// TIA Portal V20 export
VAR_GLOBAL   // PLC tag table "laser_out_macsa"
   "-XT500_output_mode" AT %QD295 : DWord;   // Pole - výber pole podle čísla max 255
   "-XT500_output_byte_1" AT %QB295 : Byte;
   "-XT500_output_byte_2" AT %QB296 : Byte;
   "-XT500_output_byte_3" AT %QB297 : Byte;
   "-XT500_output_byte_4" AT %QB298 : Byte;
   "-XT500_output_copies" AT %QD299 : DWord;
   "-XT500_output_byte_5" AT %QB299 : Byte;   // zapisovaná data
   "-XT500_output_byte_6" AT %QB300 : Byte;   // zapisovaná data
   "-XT500_output_byte_7" AT %QB301 : Byte;   // zapisovaná data
   "-XT500_output_byte_8" AT %QB302 : Byte;   // zapisovaná data
   "-XT500_output_byte_9" AT %QB303 : Byte;   // zapisovaná data
   "-XT500_output_batch" AT %QD303 : DWord;
   "-XT500_output_byte_10" AT %QB304 : Byte;   // zapisovaná data
   "-XT500_output_byte_11" AT %QB305 : Byte;   // zapisovaná data
   "-XT500_output_byte_12" AT %QB306 : Byte;   // zapisovaná data
   "-XT500_output_filename_1" AT %QB307 : Byte;   // zápid textu v asci pro volbu programu + další data
   "-XT500_output_filename_2" AT %QB308 : Byte;   // zápid textu v asci pro volbu programu + další data
   "-XT500_output_filename_3" AT %QB309 : Byte;   // zápid textu v asci pro volbu programu + další data
   "-XT500_output_filename_4" AT %QB310 : Byte;   // zápid textu v asci pro volbu programu + další data
   "-XT500_output_filename_5" AT %QB311 : Byte;   // zápid textu v asci pro volbu programu + další data
   "-XT500_output_filename_6" AT %QB312 : Byte;   // zápid textu v asci pro volbu programu + další data
   "-XT500_output_filename_7" AT %QB313 : Byte;   // zápid textu v asci pro volbu programu + další data
   "-XT500_output_filename_8" AT %QB314 : Byte;   // zápid textu v asci pro volbu programu + další data
   "-XT500_output_filename_9" AT %QB315 : Byte;   // zápid textu v asci pro volbu programu + další data
   "-XT500_output_filename_10" AT %QB316 : Byte;   // zápid textu v asci pro volbu programu + další data
   "-XT500_output_filename_11" AT %QB317 : Byte;   // zápid textu v asci pro volbu programu + další data
   "-XT500_output_filename_12" AT %QB318 : Byte;   // zápid textu v asci pro volbu programu + další data
   "-XT500_output_filename_13" AT %QB319 : Byte;   // zápid textu v asci pro volbu programu + další data
   "-XT500_output_filename_14" AT %QB320 : Byte;   // zápid textu v asci pro volbu programu + další data
   "-XT500_output_filename_15" AT %QB321 : Byte;   // zápid textu v asci pro volbu programu + další data
   "-XT500_output_filename_16" AT %QB322 : Byte;   // zápid textu v asci pro volbu programu + další data
   "-XT500_output_filename_17" AT %QB323 : Byte;   // zápid textu v asci pro volbu programu + další data
   "-XT500_command_number" AT %QB293 : Byte;   // výběr daného komandu v podobě čísla podle návodu zadavano v decu pozor na převod mezi word a int ----------- 6 zapis dat 16 vypal 1 otevření zprávy
   "-XT500_command_triger" AT %QB294 : Byte;   // 1= proveď příkaz
   "-XT500_output_filename_18" AT %QB324 : Byte;   // zápid textu v asci pro volbu programu + další data
   "-XT500_output_filename_19" AT %QB325 : Byte;   // zápid textu v asci pro volbu programu + další data
   "-XT500_output_filename_20" AT %QB326 : Byte;   // zápid textu v asci pro volbu programu + další data
   "-XT500_output_filename_21" AT %QB327 : Byte;   // zápid textu v asci pro volbu programu + další data
   "-XT500_output_filename_22" AT %QB328 : Byte;   // zápid textu v asci pro volbu programu + další data
   "-XT500_output_filename_23" AT %QB329 : Byte;   // zápid textu v asci pro volbu programu + další data
   "-XT500_output_filename_24" AT %QB330 : Byte;   // zápid textu v asci pro volbu programu + další data
   "-XT500_output_filename_25" AT %QB331 : Byte;   // zápid textu v asci pro volbu programu + další data
   "-XT500_output_filename_26" AT %QB332 : Byte;   // zápid textu v asci pro volbu programu + další data
   "-XT500_output_filename_27" AT %QB333 : Byte;   // zápid textu v asci pro volbu programu + další data
   "-XT500_output_filename_28" AT %QB334 : Byte;   // zápid textu v asci pro volbu programu + další data
   "-XT500_output_filename_29" AT %QB335 : Byte;   // zápid textu v asci pro volbu programu + další data
   "-XT500_output_filename_30" AT %QB336 : Byte;   // zápid textu v asci pro volbu programu + další data
   "-XT500_output_filename_31" AT %QB337 : Byte;   // zápid textu v asci pro volbu programu + další data
   "-XT500_output_filename_32" AT %QB338 : Byte;   // zápid textu v asci pro volbu programu + další data
   "-XT500_output_filename_33" AT %QB339 : Byte;   // zápid textu v asci pro volbu programu + další data
   "-XT500_output_filename_34" AT %QB340 : Byte;   // zápid textu v asci pro volbu programu + další data
   "-XT500_output_filename_35" AT %QB341 : Byte;   // zápid textu v asci pro volbu programu + další data
   "-XT500_output_filename_36" AT %QB342 : Byte;   // zápid textu v asci pro volbu programu + další data
   "-XT500_output_filename_37" AT %QB343 : Byte;   // zápid textu v asci pro volbu programu + další data
   "-XT500_output_filename_38" AT %QB344 : Byte;   // zápid textu v asci pro volbu programu + další data
   "-XT500_output_filename_39" AT %QB345 : Byte;   // zápid textu v asci pro volbu programu + další data
   "-XT500_output_filename_40" AT %QB346 : Byte;   // zápid textu v asci pro volbu programu + další data
   "-XT500_output_filename_41" AT %QB347 : Byte;   // zápid textu v asci pro volbu programu + další data
   "-XT500_output_filename_42" AT %QB348 : Byte;   // zápid textu v asci pro volbu programu + další data
   "-XT500_output_filename_43" AT %QB349 : Byte;   // zápid textu v asci pro volbu programu + další data
   "-XT500_output_filename_44" AT %QB350 : Byte;   // zápid textu v asci pro volbu programu + další data
   "-XT500_output_filename_45" AT %QB351 : Byte;   // zápid textu v asci pro volbu programu + další data
   "-XT500_output_filename_46" AT %QB352 : Byte;   // zápid textu v asci pro volbu programu + další data
   "-XT500_output_filename_47" AT %QB353 : Byte;   // zápid textu v asci pro volbu programu + další data
   "-XT500_output_filename_48" AT %QB354 : Byte;   // zápid textu v asci pro volbu programu + další data
   "-XT500_output_filename_49" AT %QB355 : Byte;   // zápid textu v asci pro volbu programu + další data
   "-XT500_output_filename_50" AT %QB356 : Byte;   // zápid textu v asci pro volbu programu + další data
   "-XT500_output_filename_51" AT %QB357 : Byte;   // zápid textu v asci pro volbu programu + další data
   "-XT500_output_filename_52" AT %QB358 : Byte;   // zápid textu v asci pro volbu programu + další data
   "-XT500_output_filename_53" AT %QB359 : Byte;   // zápid textu v asci pro volbu programu + další data
   "-XT500_output_filename_54" AT %QB360 : Byte;   // zápid textu v asci pro volbu programu + další data
   "-XT500_output_filename_55" AT %QB361 : Byte;   // zápid textu v asci pro volbu programu + další data
   "-XT500_output_filename_56" AT %QB362 : Byte;   // zápid textu v asci pro volbu programu + další data
   "-XT500_output_filename_57" AT %QB363 : Byte;   // zápid textu v asci pro volbu programu + další data
   "-XT500_output_filename_58" AT %QB364 : Byte;   // zápid textu v asci pro volbu programu + další data
   "-XT500_output_filename_59" AT %QB365 : Byte;   // zápid textu v asci pro volbu programu + další data
   "-XT500_output_filename_60" AT %QB366 : Byte;   // zápid textu v asci pro volbu programu + další data
   "-XT500_output_filename_61" AT %QB367 : Byte;   // zápid textu v asci pro volbu programu + další data
   "-XT500_output_filename_62" AT %QB368 : Byte;   // zápid textu v asci pro volbu programu + další data
   "-XT500_output_filename_63" AT %QB369 : Byte;   // zápid textu v asci pro volbu programu + další data
   "-XT500_output_filename_64" AT %QB370 : Byte;   // zápid textu v asci pro volbu programu + další data
   "-XT500_output_filename_65" AT %QB371 : Byte;   // zápid textu v asci pro volbu programu + další data
   "-XT500_output_filename_66" AT %QB372 : Byte;   // zápid textu v asci pro volbu programu + další data
   "-XT500_output_filename_67" AT %QB373 : Byte;   // zápid textu v asci pro volbu programu + další data
   "-XT500_output_filename_68" AT %QB374 : Byte;   // zápid textu v asci pro volbu programu + další data
   "-XT500_output_filename_69" AT %QB375 : Byte;   // zápid textu v asci pro volbu programu + další data
   "-XT500_output_filename_70" AT %QB376 : Byte;   // zápid textu v asci pro volbu programu + další data
   "-XT500_output_filename_71" AT %QB377 : Byte;   // zápid textu v asci pro volbu programu + další data
   "-XT500_output_filename_72" AT %QB378 : Byte;   // zápid textu v asci pro volbu programu + další data
   "-XT500_output_filename_73" AT %QB379 : Byte;   // zápid textu v asci pro volbu programu + další data
   "-XT500_output_filename_74" AT %QB380 : Byte;   // zápid textu v asci pro volbu programu + další data
   "-XT500_output_filename_75" AT %QB381 : Byte;   // zápid textu v asci pro volbu programu + další data
   "-XT500_output_filename_76" AT %QB382 : Byte;   // zápid textu v asci pro volbu programu + další data
   "-XT500_output_filename_77" AT %QB383 : Byte;   // zápid textu v asci pro volbu programu + další data
   "-XT500_output_filename_78" AT %QB384 : Byte;   // zápid textu v asci pro volbu programu + další data
   "-XT500_output_filename_79" AT %QB385 : Byte;   // zápid textu v asci pro volbu programu + další data
   "-XT500_output_filename_80" AT %QB386 : Byte;   // zápid textu v asci pro volbu programu + další data
   "-XT500_output_filename_81" AT %QB387 : Byte;   // zápid textu v asci pro volbu programu + další data
   "-XT500_output_filename_82" AT %QB388 : Byte;   // zápid textu v asci pro volbu programu + další data
   "-XT500_output_filename_83" AT %QB389 : Byte;   // zápid textu v asci pro volbu programu + další data
   "-XT500_output_filename_84" AT %QB390 : Byte;   // zápid textu v asci pro volbu programu + další data
   "-XT500_output_filename_85" AT %QB391 : Byte;   // zápid textu v asci pro volbu programu + další data
   "-XT500_output_filename_86" AT %QB392 : Byte;   // zápid textu v asci pro volbu programu + další data
   "-XT500_output_filename_87" AT %QB393 : Byte;   // zápid textu v asci pro volbu programu + další data
   "-XT500_output_filename_88" AT %QB394 : Byte;   // zápid textu v asci pro volbu programu + další data
   "-XT500_output_filename_89" AT %QB395 : Byte;   // zápid textu v asci pro volbu programu + další data
   "-XT500_output_filename_90" AT %QB396 : Byte;   // zápid textu v asci pro volbu programu + další data
   "-XT500_output_filename_91" AT %QB397 : Byte;   // zápid textu v asci pro volbu programu + další data
   "-XT500_output_filename_92" AT %QB398 : Byte;   // zápid textu v asci pro volbu programu + další data
   "-XT500_output_filename_93" AT %QB399 : Byte;   // zápid textu v asci pro volbu programu + další data
   "-XT500_output_filename_94" AT %QB400 : Byte;   // zápid textu v asci pro volbu programu + další data
   "-XT500_output_filename_95" AT %QB401 : Byte;   // zápid textu v asci pro volbu programu + další data
   "-XT500_output_filename_96" AT %QB402 : Byte;   // zápid textu v asci pro volbu programu + další data
   "-XT500_output_filename_97" AT %QB403 : Byte;   // zápid textu v asci pro volbu programu + další data
   "-XT500_output_filename_98" AT %QB404 : Byte;   // zápid textu v asci pro volbu programu + další data
   "-XT500_output_filename_99" AT %QB405 : Byte;   // zápid textu v asci pro volbu programu + další data
   "-XT500_output_filename_100" AT %QB406 : Byte;   // zápid textu v asci pro volbu programu + další data
   "-XT500_output_filename_101" AT %QB407 : Byte;   // zápid textu v asci pro volbu programu + další data
   "-XT500_output_filename_102" AT %QB408 : Byte;   // zápid textu v asci pro volbu programu + další data
   "-XT500_output_filename_103" AT %QB409 : Byte;   // zápid textu v asci pro volbu programu + další data
   "-XT500_output_filename_104" AT %QB410 : Byte;   // zápid textu v asci pro volbu programu + další data
   "-XT500_output_filename_105" AT %QB422 : Byte;   // zápid textu v asci pro volbu programu + další data
   "-XT500_output_filename_106" AT %QB423 : Byte;   // zápid textu v asci pro volbu programu + další data
   "-XT500_output_filename_107" AT %QB424 : Byte;   // zápid textu v asci pro volbu programu + další data
   "-XT500_output_filename_108" AT %QB425 : Byte;   // zápid textu v asci pro volbu programu + další data
   "-XT500_output_filename_109" AT %QB426 : Byte;   // zápid textu v asci pro volbu programu + další data
   "-XT500_output_filename_110" AT %QB427 : Byte;   // zápid textu v asci pro volbu programu + další data
   "-XT500_output_filename_111" AT %QB428 : Byte;   // zápid textu v asci pro volbu programu + další data
   "-XT500_output_filename_112" AT %QB429 : Byte;   // zápid textu v asci pro volbu programu + další data
   "-XT500_output_filename_113" AT %QB430 : Byte;   // zápid textu v asci pro volbu programu + další data
   "-XT500_output_filename_114" AT %QB431 : Byte;   // zápid textu v asci pro volbu programu + další data
   "-XT500_output_filename_115" AT %QB432 : Byte;   // zápid textu v asci pro volbu programu + další data
   "-XT500_output_filename_116" AT %QB433 : Byte;   // zápid textu v asci pro volbu programu + další data
   "-XT500_output_filename_117" AT %QB434 : Byte;   // zápid textu v asci pro volbu programu + další data
   "-XT500_output_filename_118" AT %QB435 : Byte;   // zápid textu v asci pro volbu programu + další data
   "-XT500_output_filename_119" AT %QB436 : Byte;   // zápid textu v asci pro volbu programu + další data
   "-XT500_output_filename_120" AT %QB437 : Byte;   // zápid textu v asci pro volbu programu + další data
   "-XT500_output_filename_121" AT %QB438 : Byte;   // zápid textu v asci pro volbu programu + další data
   "-XT500_output_filename_122" AT %QB439 : Byte;   // zápid textu v asci pro volbu programu + další data
   "-XT500_output_filename_123" AT %QB440 : Byte;   // zápid textu v asci pro volbu programu + další data
   "-XT500_output_filename_124" AT %QB441 : Byte;   // zápid textu v asci pro volbu programu + další data
   "-XT500_output_filename_125" AT %QB442 : Byte;   // zápid textu v asci pro volbu programu + další data
   "-XT500_output_filename_126" AT %QB443 : Byte;   // zápid textu v asci pro volbu programu + další data
   "-XT500_output_filename_127" AT %QB444 : Byte;   // zápid textu v asci pro volbu programu + další data
   "-XT500_output_filename_128" AT %QB445 : Byte;   // zápid textu v asci pro volbu programu + další data
   "-XT500_output_filename_129" AT %QB446 : Byte;   // zápid textu v asci pro volbu programu + další data
   "-XT500_output_filename_130" AT %QB447 : Byte;   // zápid textu v asci pro volbu programu + další data
   "-XT500_output_filename_131" AT %QB448 : Byte;   // zápid textu v asci pro volbu programu + další data
   "-XT500_output_filename_132" AT %QB449 : Byte;   // zápid textu v asci pro volbu programu + další data
   "-XT500_output_filename_133" AT %QB450 : Byte;   // zápid textu v asci pro volbu programu + další data
   "-XT500_output_filename_134" AT %QB451 : Byte;   // zápid textu v asci pro volbu programu + další data
   "-XT500_output_filename_135" AT %QB452 : Byte;   // zápid textu v asci pro volbu programu + další data
   "-XT500_output_filename_136" AT %QB453 : Byte;   // zápid textu v asci pro volbu programu + další data
   "-XT500_output_filename_137" AT %QB454 : Byte;   // zápid textu v asci pro volbu programu + další data
   "-XT500_output_filename_138" AT %QB455 : Byte;   // zápid textu v asci pro volbu programu + další data
END_VAR
